(* IEC 61131-3 sources: volt/packages/volt-lsp-iec/test-corpus/twincat-project14/TwinCAT Project14/PLC/Untitled2/Untitled2 Project/References/Tc3_Module, 38 files *)

(* ---- Global_Version.gvl ---- *)
VAR_GLOBAL
	stLibVersion_Tc3_Module : ST_LibVersion;
END_VAR

(* ---- GVL.gvl ---- *)
VAR_GLOBAL
	S_OK : HRESULT;
	S_FALSE : HRESULT;
	S_PENDING : HRESULT;
	S_WATCHDOG_TIMEOUT : HRESULT;
	E_FAIL : HRESULT;
	ERR_INVALID_PARAM : HRESULT;
	OTCID_CreateNewId : OTCID;
	OTCID_FirstFreeId : OTCID;
	OTCID_LastFreeId : OTCID;
	NULL : PVOID;
END_VAR

(* ---- ExCpHndFunc.pou ---- *)
FUNCTION ExCpHndFunc : UDINT
VAR_INPUT
	pUsr : PVOID;
	pExcpHndPara : PVOID;
END_VAR
END_FUNCTION

(* ---- F_CPUCounter.pou ---- *)
FUNCTION F_CPUCounter : BOOL
VAR_INPUT
	counter : ULINT;
END_VAR
END_FUNCTION

(* ---- F_TcLicSrv_TakeLicense.pou ---- *)
FUNCTION F_TcLicSrv_TakeLicense : HRESULT
VAR_INPUT
	refLicenseId : REFERENCE TO GUID;
END_VAR
END_FUNCTION

(* ---- FAILED.pou ---- *)
FUNCTION FAILED : BOOL
VAR_INPUT
	hr : HRESULT;
END_VAR
END_FUNCTION

(* ---- FW_GetAppState.pou ---- *)
FUNCTION FW_GetAppState : UDINT
END_FUNCTION

(* ---- FW_MemCmp.pou ---- *)
FUNCTION FW_MemCmp : DINT
VAR_INPUT
	pBuf1 : PVOID;
	pBuf2 : PVOID;
	cbLen : UDINT;
END_VAR
END_FUNCTION

(* ---- FW_MemCpy.pou ---- *)
FUNCTION FW_MemCpy : UDINT
VAR_INPUT
	pDest : PVOID;
	pSrc : PVOID;
	cbLen : UDINT;
END_VAR
END_FUNCTION

(* ---- FW_MemSet.pou ---- *)
FUNCTION FW_MemSet : UDINT
VAR_INPUT
	pDest : PVOID;
	nFillByte : USINT;
	cbLen : UDINT;
END_VAR
END_FUNCTION

(* ---- FW_ObjMgr_CreateAndInitInstance.pou ---- *)
FUNCTION FW_ObjMgr_CreateAndInitInstance : HRESULT
VAR_INPUT
	clsId : CLSID;
	iid : IID;
	pipUnk : POINTER TO ITcUnknown;
	objId : UDINT;
	parentId : UDINT;
	name : REFERENCE TO STRING;
	state : UDINT;
	pInitData : POINTER TO TComInitDataHdr;
END_VAR
END_FUNCTION

(* ---- FW_ObjMgr_CreateInstance.pou ---- *)
FUNCTION FW_ObjMgr_CreateInstance : HRESULT
VAR_INPUT
	clsId : CLSID;
	iid : IID;
	pipUnk : POINTER TO ITcUnknown;
END_VAR
END_FUNCTION

(* ---- FW_ObjMgr_DeleteInstance.pou ---- *)
FUNCTION FW_ObjMgr_DeleteInstance : HRESULT
VAR_INPUT
	pipUnk : POINTER TO ITcUnknown;
END_VAR
END_FUNCTION

(* ---- FW_ObjMgr_DeregisterObject.pou ---- *)
FUNCTION FW_ObjMgr_DeregisterObject : HRESULT
VAR_INPUT
	oidApp : OTCID;
	oidObj : OTCID;
	bInCopyCode : BOOL;
END_VAR
END_FUNCTION

(* ---- FW_ObjMgr_GetObjectInstance.pou ---- *)
FUNCTION FW_ObjMgr_GetObjectInstance : HRESULT
VAR_INPUT
	oid : OTCID;
	iid : IID;
	pipUnk : POINTER TO ITcUnknown;
END_VAR
END_FUNCTION

(* ---- FW_ObjMgr_GetObjectServer.pou ---- *)
FUNCTION FW_ObjMgr_GetObjectServer : HRESULT
VAR_INPUT
	oidApp : OTCID;
	pipSrv : POINTER TO ITComObjectServer;
END_VAR
END_FUNCTION

(* ---- FW_ObjMgr_RegisterObject.pou ---- *)
FUNCTION FW_ObjMgr_RegisterObject : HRESULT
VAR_INPUT
	oidApp : OTCID;
	oidObj : OTCID;
	bInCopyCode : BOOL;
	ipUnk : ITcUnknown;
END_VAR
END_FUNCTION

(* ---- FW_SafeRelease.pou ---- *)
FUNCTION FW_SafeRelease : HRESULT
VAR_INPUT
	pipUnk : POINTER TO ITcUnknown;
END_VAR
END_FUNCTION

(* ---- Fw_Trace.pou ---- *)
FUNCTION Fw_Trace : DINT
VAR_INPUT
	val : DINT;
	text : STRING(255);
END_VAR
END_FUNCTION

(* ---- GuidsEqual.pou ---- *)
FUNCTION GuidsEqual : BOOL
VAR_INPUT
	pGuidA : POINTER TO GUID;
	pGuidB : POINTER TO GUID;
END_VAR
END_FUNCTION

(* ---- ITCUNKNOWN_TO_PVOID.pou ---- *)
FUNCTION ITCUNKNOWN_TO_PVOID : PVOID
VAR_INPUT
	itcUnknown : ITcUnknown;
END_VAR
END_FUNCTION

(* ---- MEMCMP.pou ---- *)
FUNCTION MEMCMP : DINT
VAR_INPUT
	pBuf1 : PVOID;
	pBuf2 : PVOID;
	n : UDINT;
END_VAR
END_FUNCTION

(* ---- MEMCPY.pou ---- *)
FUNCTION MEMCPY : UDINT
VAR_INPUT
	destAddr : PVOID;
	srcAddr : PVOID;
	n : UDINT;
END_VAR
END_FUNCTION

(* ---- MEMSET.pou ---- *)
FUNCTION MEMSET : UDINT
VAR_INPUT
	destAddr : PVOID;
	fillByte : USINT;
	n : UDINT;
END_VAR
END_FUNCTION

(* ---- POINTERTOINTERFACE_TO_PVOID.pou ---- *)
FUNCTION POINTERTOINTERFACE_TO_PVOID : PVOID
VAR_INPUT
	pTmp : POINTER TO PVOID;
END_VAR
END_FUNCTION

(* ---- PTComInitDataElmHdrDATA.pou ---- *)
FUNCTION PTComInitDataElmHdrDATA : POINTER TO TComInitDataElmHdr
VAR_INPUT
	pTComInitDataElmHdr : POINTER TO TComInitDataElmHdr;
END_VAR
END_FUNCTION

(* ---- PTComInitDataElmHdrNEXTHDR.pou ---- *)
FUNCTION PTComInitDataElmHdrNEXTHDR : POINTER TO TComInitDataElmHdr
VAR_INPUT
	pTComInitDataElmHdr : POINTER TO TComInitDataElmHdr;
END_VAR
END_FUNCTION

(* ---- PTComInitDataElmHdrSIZEOF.pou ---- *)
FUNCTION PTComInitDataElmHdrSIZEOF : DINT
VAR_INPUT
	pTComInitDataElmHdr : POINTER TO TComInitDataElmHdr;
END_VAR
END_FUNCTION

(* ---- PVOID_TO_ITCUNKNOWN.pou ---- *)
FUNCTION PVOID_TO_ITCUNKNOWN : ITcUnknown
VAR_INPUT
	pVoid : PVOID;
END_VAR
END_FUNCTION

(* ---- PVOID_TO_POINTERTOINTERFACE.pou ---- *)
FUNCTION PVOID_TO_POINTERTOINTERFACE : POINTER TO ITcUnknown
VAR_INPUT
	pVoid : PVOID;
END_VAR
END_FUNCTION

(* ---- SizeOfCString.pou ---- *)
FUNCTION SizeOfCString : UDINT
VAR_INPUT
	myCString : POINTER TO STRING;
END_VAR
END_FUNCTION

(* ---- SUCCEEDED.pou ---- *)
FUNCTION SUCCEEDED : BOOL
VAR_INPUT
	hr : HRESULT;
END_VAR
END_FUNCTION

(* ---- TaskFnc.pou ---- *)
FUNCTION TaskFnc : UDINT
VAR_INPUT
	pUsr : PVOID;
END_VAR
END_FUNCTION

(* ---- IecTaskModule.pou ---- *)
FUNCTION_BLOCK IecTaskModule
END_FUNCTION_BLOCK

(* ---- IecTaskModulePost.pou ---- *)
FUNCTION_BLOCK IecTaskModulePost
END_FUNCTION_BLOCK

(* ---- TcBaseModule.pou ---- *)
FUNCTION_BLOCK TcBaseModule
END_FUNCTION_BLOCK

(* ---- TcBaseModuleRegistered.pou ---- *)
FUNCTION_BLOCK TcBaseModuleRegistered
END_FUNCTION_BLOCK

(* ---- TcBaseModuleRegistered2.pou ---- *)
FUNCTION_BLOCK TcBaseModuleRegistered2
VAR_OUTPUT
	objID : OTCID;
END_VAR
END_FUNCTION_BLOCK
